{attribute 'no_assign'}
FUNCTION_BLOCK FB_LN_WTURBINE_LD0_WTUR1 EXTENDS FB_AcsiCommonLogicalNodeClass
VAR_INPUT
	Beh: FB_DO_WTURBINE_LD0_WTUR1_Beh := (sClass:='ENS', bLinkResult:=THIS^.AddDataToContainer(ipData:=Beh));
	TotWh: FB_DO_WTURBINE_LD0_WTUR1_TotWh := (sClass:='CTE', bLinkResult:=THIS^.AddDataToContainer(ipData:=TotWh));
	TurSt: FB_DO_WTURBINE_LD0_WTUR1_TurSt := (sClass:='STV', bLinkResult:=THIS^.AddDataToContainer(ipData:=TurSt));
	W: FB_DO_WTURBINE_LD0_WTUR1_W := (sClass:='MV', bLinkResult:=THIS^.AddDataToContainer(ipData:=W));
	TurOp: FB_DO_WTURBINE_LD0_WTUR1_TurOp := (sClass:='CMD', bLinkResult:=THIS^.AddDataToContainer(ipData:=TurOp));
	DmdWSpt: FB_DO_WTURBINE_LD0_WTUR1_DmdWSpt := (sClass:='SPV', bLinkResult:=THIS^.AddDataToContainer(ipData:=DmdWSpt));
	TurCtl: FB_DO_WTURBINE_LD0_WTUR1_TurCtl := (sClass:='CMD', bLinkResult:=THIS^.AddDataToContainer(ipData:=TurCtl));
END_VAR
VAR
END_VAR

END_FUNCTION_BLOCK

(* stored: Version 1.1.0.1
   POU FB_LN_WTURBINE_LD0_WTUR1: Id {4c88211b-29d2-4499-89b9-726757d83e70}, SpecialFunc None *)
